ABB RAPID module: JointTargets.prg

%%%
  VERSION:1
  LANGUAGE:ENGLISH
%%%
MODULE MOD_JointTargets

    ! -------------------------------
    ! Define customized variables here
    ! ...

	! Tool variables:
	PERS tooldata Tool1 := [TRUE,[[10.000,0.000,120.000],[0.99144486,0.00000000,0.13052619,0.00000001]],[1,[0,0,20],[1,0,0,0],0,0,0.005]];

	! Reference variables:
	PERS wobjdata Frame2 := [FALSE, TRUE, "", [[100.000,-50.000,20.000],[0.96592583,0.00000000,0.00000000,0.25881905]],[[0,0,0],[1,0,0,0]]];

	PROC Main()
		ConfJ \On;
		ConfL \Off;
		! Program generated by VerticalBot Studio for ABB IRB 120-3/0.6 on 25/10/2026 12:00:00
		! Using nominal kinematics.
		MoveAbsJ [[-10.000000,10.000000,20.000000,30.000000,40.000000,-50.000000],[9E+09,9E+09,9E+09,9E+09,9E+09,9E+09]],v500,z1,Tool1 \WObj:=Frame2;
		MoveL CalcRobT([[-2.000000,14.000000,20.000000,30.000000,40.000000,-50.000000],[9E+09,9E+09,9E+09,9E+09,9E+09,9E+09]],Tool1 \WObj:=Frame2),v500,z1,Tool1 \WObj:=Frame2;
		MoveAbsJ [[-2.000000,14.000000,20.000000,30.000000,40.000000,-50.000000],[9E+09,9E+09,9E+09,9E+09,9E+09,9E+09]],v500,z1,Tool1 \WObj:=Frame2;
		MoveL [[289.255,-125.996,274.474],[0.13100243,0.07930186,0.98767984,0.03221959],[-1,0,-1,0],[9E+09,9E+09,9E+09,9E+09,9E+09,9E+09]],v500,z1,Tool1 \WObj:=Frame2;
		MoveL CalcRobT([[-2.000000,14.000000,20.000000,30.000000,40.000000,-50.000000],[9E+09,9E+09,9E+09,9E+09,9E+09,9E+09]],Tool1 \WObj:=Frame2),v500,z1,Tool1 \WObj:=Frame2;
		MoveAbsJ [[-10.000000,10.000000,20.000000,30.000000,40.000000,-50.000000],[9E+09,9E+09,9E+09,9E+09,9E+09,9E+09]],v500,z5,Tool1 \WObj:=Frame2;
		MoveL CalcRobT([[-2.000000,14.000000,20.000000,30.000000,40.000000,-50.000000],[9E+09,9E+09,9E+09,9E+09,9E+09,9E+09]],Tool1 \WObj:=Frame2),v500,z5,Tool1 \WObj:=Frame2;
		MoveAbsJ [[-2.000000,14.000000,20.000000,30.000000,40.000000,-50.000000],[9E+09,9E+09,9E+09,9E+09,9E+09,9E+09]],v500,z5,Tool1 \WObj:=Frame2;
		MoveL [[289.255,-125.996,274.474],[0.13100243,0.07930186,0.98767984,0.03221959],[-1,0,-1,0],[9E+09,9E+09,9E+09,9E+09,9E+09,9E+09]],v500,z5,Tool1 \WObj:=Frame2;
		MoveL CalcRobT([[-2.000000,14.000000,20.000000,30.000000,40.000000,-50.000000],[9E+09,9E+09,9E+09,9E+09,9E+09,9E+09]],Tool1 \WObj:=Frame2),v500,z5,Tool1 \WObj:=Frame2;
		MoveAbsJ [[-10.000000,10.000000,20.000000,30.000000,40.000000,-50.000000],[9E+09,9E+09,9E+09,9E+09,9E+09,9E+09]],v500,fine,Tool1 \WObj:=Frame2;
	ENDPROC

ENDMODULE
